(* IEC 61131-3 sources: Lasal-MCP/examples/SampleSource/LASALScreenAdvancedSolution/LASALScreenAdvancedSolution/LASALScreenAdvacnedSolution/Stations/Terminal/HMI/Class/FileHandling, 1 file *)

(* ---- FileHandling.st ---- *)
(*!
<Class
	Name               = "FileHandling"
	Revision           = "0.0"
	RealtimeTask       = "false"
	CyclicTask         = "false"
	BackgroundTask     = "true"
	DefBackground      = "50 ms"
	Sigmatek           = "false"
	OSInterface        = "false"
	HighPriority       = "false"
	Automatic          = "false"
	UpdateMode         = "Prescan"
	SharedCommandTable = "true"
	Objectsize         = "(720,180)">
	<Channels>
		<Server Name="DriveName1" Visualized="true" Remotely="true" Initialize="true" WriteProtected="false" Retentive="false"/>
		<Server Name="FileExtension1" Visualized="true" Remotely="true" Initialize="true" WriteProtected="false" Retentive="false"/>
		<Server Name="FileIsCreated" Visualized="false" Initialize="false" WriteProtected="true" Retentive="false"/>
		<Server Name="FileName1" Visualized="true" Remotely="true" Initialize="true" WriteProtected="false" Retentive="false"/>
		<Server Name="IntError" Visualized="false" Initialize="false" WriteProtected="true" Retentive="false"/>
		<Server Name="StartFileWrite" Visualized="false" Initialize="false" WriteProtected="false" Retentive="false"/>
		<Server Name="Steps" Visualized="false" Initialize="false" WriteProtected="true" Retentive="false"/>
		<Client Name="_FileSys" Required="false" Internal="false"/>
		<Client Name="_StdLib" Required="false" Internal="false"/>
		<Client Name="DriveName" Required="true" Internal="true"/>
		<Client Name="FileExtension" Required="true" Internal="true"/>
		<Client Name="FileName" Required="true" Internal="true"/>
		<Client Name="FileRead" Required="true" Internal="false"/>
		<Client Name="SigCLib" Required="false" Internal="false"/>
	</Channels>
	<Network Name="FileHandling">
		<!-- List of Components in this network -->
		<Components>
			<Object
				Name       = "DriveName"
				Class      = "StringRAM"
				Position   = "(60,390)"
				Visualized = "true"
				Remotely   = "true">
				<Channels>
					<Server Name="Data"/>
					<Client Name="SingleRealloc" Value="1"/>
					<Client Name="UseFile"/>
				</Channels>
			</Object>
			<Object
				Name       = "FileExtension"
				Class      = "StringRAM"
				Position   = "(60,810)"
				Visualized = "true"
				Remotely   = "true">
				<Channels>
					<Server Name="Data"/>
					<Client Name="SingleRealloc" Value="1"/>
					<Client Name="UseFile"/>
				</Channels>
			</Object>
			<Object
				Name       = "FileName"
				Class      = "StringRAM"
				Position   = "(60,600)"
				Visualized = "true"
				Remotely   = "true">
				<Channels>
					<Server Name="Data"/>
					<Client Name="SingleRealloc" Value="1"/>
					<Client Name="UseFile"/>
				</Channels>
			</Object>
		</Components>
		<Comments>
		</Comments>
		<!-- List of Connections in this network -->
		<Connections>
			<Connection Source="this.DriveName" Destination="DriveName.Data"/>
			<Connection Source="this.FileName" Destination="FileName.Data"/>
			<Connection Source="this.FileExtension" Destination="FileExtension.Data"/>
			<Connection Source="this.DriveName1" Destination="DriveName.Data" Vertices="(728,450),(556,480),"/>
			<Connection Source="this.FileName1" Destination="FileName.Data" Vertices="(728,510),(556,690),"/>
			<Connection Source="this.FileExtension1" Destination="FileExtension.Data" Vertices="(728,570),(556,900),"/>
		</Connections>
		<!-- Headerfiles -->
		<Options>
		</Options>
	</Network>
</Class>
*)
FileHandling : CLASS
	TYPE
	  t_e_FILE_STEPS :  //! <Type Public="true" Name="t_e_FILE_STEPS"/>
	  (
	    tFH_Idle,
	    tFH_FileCreate,
	    tFH_WaitFileCreated,
	    tFH_FileClose,
	    tFH_WaitFileClosed,
	    tFH_FileOpen,
	    tFH_WaitFileOpened,
	    tFH_FileWrite,
	    tFH_WaitFileWritten,
	    tFH_FileRead,
	    tFH_WaitFileRead,
	    tFH_Error
	  )$UDINT;
	END_TYPE
  //Servers:
	Steps 	: SvrChCmd_t_e_FILE_STEPS_PTofCls_FileHandling;
	StartFileWrite 	: SvrCh_DINT;
	FileIsCreated 	: SvrCh_DINT;
	IntError 	: SvrCh_DINT;
	DriveName1 	: SvrCh_UDINT;
	FileName1 	: SvrCh_UDINT;
	FileExtension1 	: SvrCh_UDINT;
  //Clients:
	_FileSys 	: CltChCmd__FileSys;
	SigCLib 	: CltChCmd_SigCLib;
	DriveName 	: CltChCmd_StringRAM;
	FileName 	: CltChCmd_StringRAM;
	FileExtension 	: CltChCmd_StringRAM;
	_StdLib 	: CltChCmd__StdLib;
	FileRead 	: CltChCmd_FileRead;
  //Variables:
		FullFileName : ARRAY [0..255] OF CHAR;

		StringLength 	: UDINT;
		pError 	: ^CHAR;
		FileHandle 	: DINT;
		FileWritten 	: DINT;
		FunctionID 	: DINT;
		FunctionState 	: DINT;
		Length 	: UDINT;
		pSaveData 	: ^DINT;
		ReadFile 	: BOOL;
  //Functions:

	FUNCTION VIRTUAL GLOBAL Init;

	FUNCTION VIRTUAL GLOBAL Background
		VAR_INPUT
			EAX 	: UDINT;
		END_VAR
		VAR_OUTPUT
			state (EAX) 	: UDINT;
		END_VAR;

	FUNCTION GLOBAL StartWrite
		VAR_INPUT
			pData 	: ^DINT;
			Amount 	: UDINT;
		END_VAR
		VAR_OUTPUT
			Retcode 	: DINT;
		END_VAR;

	FUNCTION VIRTUAL GLOBAL DriveName1::Read
		VAR_OUTPUT
			output (EAX) 	: UDINT;
		END_VAR;

	FUNCTION VIRTUAL GLOBAL DriveName1::Write
		VAR_INPUT
			input (EAX) 	: UDINT;
		END_VAR
		VAR_OUTPUT
			result (EAX) 	: UDINT;
		END_VAR;

	FUNCTION VIRTUAL GLOBAL FileName1::Read
		VAR_OUTPUT
			output (EAX) 	: UDINT;
		END_VAR;

	FUNCTION VIRTUAL GLOBAL FileName1::Write
		VAR_INPUT
			input (EAX) 	: UDINT;
		END_VAR
		VAR_OUTPUT
			result (EAX) 	: UDINT;
		END_VAR;

	FUNCTION VIRTUAL GLOBAL FileExtension1::Read
		VAR_OUTPUT
			output (EAX) 	: UDINT;
		END_VAR;

	FUNCTION VIRTUAL GLOBAL FileExtension1::Write
		VAR_INPUT
			input (EAX) 	: UDINT;
		END_VAR
		VAR_OUTPUT
			result (EAX) 	: UDINT;
		END_VAR;
  //Tables:
	FUNCTION @STD
		VAR_OUTPUT
			ret_code	: CONFSTATES;
		END_VAR;
	FUNCTION GLOBAL TAB @CT_;
END_CLASS;

#pragma using StringRAM
#pragma usingLtd _FileSys
#pragma usingLtd _StdLib
#pragma usingLtd FileRead
#pragma usingLtd SigCLib

FUNCTION VIRTUAL GLOBAL FileHandling::Init

  if (_FirstScan = TRUE) then
    Steps := tFH_FileCreate; // Create file in the beginning
  end_if;

END_FUNCTION

FUNCTION VIRTUAL GLOBAL FileHandling::Background
	VAR_INPUT
		EAX 	: UDINT;
	END_VAR
	VAR_OUTPUT
		state (EAX) 	: UDINT;
	END_VAR
  VAR
    Temp : ARRAY[0..255] of CHAR;
    retCode : UDINT;
  END_VAR

  //******************************************************************
  //  File Handling
  //******************************************************************
  case Steps of
  //******************************************************************
  	tFH_Idle:
      if (StartFileWrite = 1) then
        StartFileWrite := 0;
        Steps := tFH_FileOpen;
      end_if;

  //******************************************************************
  	tFH_FileCreate:
      // ==========  get drive name  ==========
      retCode := DriveName.TxtGet(pdst:= #Temp[0],
                                        dstsize:= sizeof(Temp));

      if (retCode = 0) then

        intError := -1;
        Steps := tFH_Error;
        return;

      end_if;

      pError := SigCLib.StrCpy(dst0:= #FullFileName[0],
                               src0:= #Temp[0]);

      if (pError <> #FullFileName[0]) then
        IntError := -2;
        Steps := tFH_Error;
        return;
      end_if;

      // ==========  get file name  ==========
      retCode := FileName.TxtGet(pdst:= #Temp[0],
                                        dstsize:= sizeof(Temp));

      if (retCode = 0) then

        intError := -3;
        Steps := tFH_Error;
        return;

      end_if;

      pError := SigCLib.StrCat(ps1:= #FullFileName[0],
                               ps2:= #Temp[0]);

      if (pError <> #FullFileName[0]) then
        IntError := -4;
        Steps := tFH_Error;
        return;
      end_if;

      // ==========  get file extension  ==========
      retCode := FileExtension.TxtGet(pdst:= #Temp[0],
                                       dstsize:= sizeof(Temp));

      if (retCode = 0) then

        intError := -5;
        Steps := tFH_Error;
        return;

      end_if;

      pError := SigCLib.StrCat(ps1:= #FullFileName[0],
                               ps2:= #Temp[0]);

      if (pError <> #FullFileName[0]) then
        IntError := -6;
        Steps := tFH_Error;
        return;
      end_if;

      FunctionID := _FileSys.FileCreate_A(Async:= 1,
                                          dpne:= #FullFileName[0],
                                          size:= 1 MB,
                                          fill:= 0,
                                          att:= ATT_CREATE_ALWAYS);

      Steps := tFH_WaitFileCreated;

  //******************************************************************
  	tFH_WaitFileCreated:

      FunctionState := _FileSys.GetAsyncState(ID:= to_udint(FunctionID),
                                              Erg:= #FileHandle);

      case FunctionState of
        //-----------------------------------
        0:
          if (FileHandle >= 0) then
            Steps := tFH_FileClose;
            FileIsCreated := 1;
          else
            IntError := -7;
            Steps := tFH_Error;
          end_if;

        //-----------------------------------
        RT_ERG_DELETED,
        RT_INVALID_ID:
          IntError := -8;
          Steps := tFH_Error;

        //-----------------------------------
        RT_NOT_STARTED,
        RT_IN_PROGRESS:

      end_case;

  //******************************************************************
  	tFH_FileClose:

      FunctionID := _FileSys.FileClose_A(Async:= 1,
                                         handle:= FileHandle);

      Steps := tFH_WaitFileClosed;

  //******************************************************************
  	tFH_WaitFileClosed:

      FunctionState := _FileSys.GetAsyncState(ID:= to_udint(FunctionID),
                                              Erg:= #FileHandle);

      case FunctionState of
        //-----------------------------------
        0:
          if (FileHandle >= 0) then

            if (FileIsCreated = 1) then
              Steps := tFH_Idle;
            end_if;

          else
            IntError := -9;
            Steps := tFH_Error;
          end_if;

        //-----------------------------------
        RT_ERG_DELETED,
        RT_INVALID_ID:
          IntError := -10;
          Steps := tFH_Error;

        //-----------------------------------
        RT_NOT_STARTED,
        RT_IN_PROGRESS:

      end_case;

  //******************************************************************
  	tFH_FileOpen:

      FunctionID := _FileSys.FileOpen_A(Async:= 1,
                                        filename:= #FullFileName[0],
                                        attributes:= ATT_READ_WRITE);

      Steps := tFH_WaitFileOpened;

  //******************************************************************
  	tFH_WaitFileOpened:

      FunctionState := _FileSys.GetAsyncState(ID:= to_udint(FunctionID),
                                              Erg:= #FileHandle);

      case FunctionState of
        //-----------------------------------
        0:
          if (FileHandle >= 0) then

            Steps := tFH_FileWrite;

          elsif (FileHandle = -16) then
            Steps := tFH_FileCreate;
          else
            IntError := -11;
            Steps := tFH_Error;
          end_if;

        //-----------------------------------
        RT_ERG_DELETED,
        RT_INVALID_ID:
          IntError := -12;
          Steps := tFH_Error;

        //-----------------------------------
        RT_NOT_STARTED,
        RT_IN_PROGRESS:

      end_case;

  //******************************************************************
  	tFH_FileWrite:

      FunctionID := _FileSys.FileWrite_A(Async:= 1,
                                         handle:= FileHandle,
                                         buffer:= pSaveData,
                                         Length:= Length);

      Steps := tFH_WaitFileWritten;

  //******************************************************************
  	tFH_WaitFileWritten:

      FunctionState := _FileSys.GetAsyncState(ID:=to_udint(FunctionID),
                                                 Erg:=#FileWritten);

      case FunctionState of
        //-----------------------------------
        0:
          if (FileWritten >= 0) then
            Steps := tFH_FileClose;
          else
            IntError := -13;
            Steps := tFH_Error;
          end_if;

        //-----------------------------------
        RT_ERG_DELETED,
        RT_INVALID_ID:
          IntError := -14;
          Steps := tFH_Error;

        //-----------------------------------
        RT_NOT_STARTED,
        RT_IN_PROGRESS:

      end_case;

  //******************************************************************
    tFH_Error:

  end_case;
  //******************************************************************
  //  End File Handling
  //******************************************************************

	state := READY;

END_FUNCTION

FUNCTION GLOBAL FileHandling::StartWrite
	VAR_INPUT
		pData 	: ^DINT;
		Amount 	: UDINT;
	END_VAR
	VAR_OUTPUT
		Retcode 	: DINT;
	END_VAR

  if (pData = NIL) then
    IntError := -14;
    Retcode := -1;
    return;
  end_if;

  if (FileIsCreated = 0) then
    Retcode := -2;
    return;
  end_if;

  pSaveData := pData;
  Length := Amount;
  ReadFile := FALSE;
  Steps := tFH_FileOpen;

END_FUNCTION

FUNCTION VIRTUAL GLOBAL FileHandling::DriveName1::Read
	VAR_OUTPUT
		output (EAX) 	: UDINT;
	END_VAR

	DriveName1 := DriveName.Data.Read();
	output := DriveName1;

END_FUNCTION

FUNCTION VIRTUAL GLOBAL FileHandling::DriveName1::Write
	VAR_INPUT
		input (EAX) 	: UDINT;
	END_VAR
	VAR_OUTPUT
		result (EAX) 	: UDINT;
	END_VAR

	DriveName1 := input;
	result := (DriveName.Data.Write(DriveName1))$UDINT;

END_FUNCTION

FUNCTION VIRTUAL GLOBAL FileHandling::FileName1::Read
	VAR_OUTPUT
		output (EAX) 	: UDINT;
	END_VAR

	FileName1 := FileName.Data.Read();
	output := FileName1;

END_FUNCTION

FUNCTION VIRTUAL GLOBAL FileHandling::FileName1::Write
	VAR_INPUT
		input (EAX) 	: UDINT;
	END_VAR
	VAR_OUTPUT
		result (EAX) 	: UDINT;
	END_VAR

	FileName1 := input;
	result := (FileName.Data.Write(FileName1))$UDINT;

END_FUNCTION

FUNCTION VIRTUAL GLOBAL FileHandling::FileExtension1::Read
	VAR_OUTPUT
		output (EAX) 	: UDINT;
	END_VAR

	FileExtension1 := FileExtension.Data.Read();
	output := FileExtension1;

END_FUNCTION

FUNCTION VIRTUAL GLOBAL FileHandling::FileExtension1::Write
	VAR_INPUT
		input (EAX) 	: UDINT;
	END_VAR
	VAR_OUTPUT
		result (EAX) 	: UDINT;
	END_VAR

	FileExtension1 := input;
	result := (FileExtension.Data.Write(FileExtension1))$UDINT;

END_FUNCTION
